Fanuc KAREL source: kt00708.KL

-- PROVISIONAL review KL for V770-1; original PC SHA256 b51188e6a006aecd14a432b9cd2e175cfca6e49dae70c71884a15528c6d5e794
-- Incomplete behavior may be omitted. Consult companion uncertainty JSON. Do not deploy.
PROGRAM KT00708
%NOLOCKGROUP
VAR
  R1 : REAL
  R2 : REAL
  OUT : BOOLEAN
BEGIN
  -- UNRESOLVED_PC offsets 5-16; opcodes 2E,23
  -- UNRESOLVED_PC offsets 21-32; opcodes 2E,23
  -- UNRESOLVED_PC offsets 37-48; opcodes 2E,23
  -- UNRESOLVED_PC offsets 53-64; opcodes 2E,23
  -- UNRESOLVED_PC offsets 69-84; opcodes 22,63,23
  -- UNRESOLVED_PC offsets 89-93; opcodes 7F
END KT00708
